Staubli VAL3: ForceData.pjx

--- ForceData.pjx ---
Parameters version=s8.15.3Cs9_BS3337 stackSize=5000 millimeterUnit=true
Data file=ForceData.dtx
Type name=tForce4Item path=Disk://LibTorque/template/Force4Item/Force4Item.pjx
Type name=tForce6Item path=Disk://LibTorque/template/Force6Item/Force6Item.pjx

--- ForceData.dtx ---
public tForce4Item tArm4Force{}
  [tp_80]
    num nMaxJnt4Force[4]
      [0] = 1029
      [1] = 254
      [2] = 833
      [3] = 15.2
    string sArmType
  [ts2_100]
    num nMaxJnt4Force[4]
      [0] = 570
      [1] = 255
      [2] = 789
      [3] = 15.6
    string sArmType
  [ts2_40]
    num nMaxJnt4Force[4]
      [0] = 570
      [1] = 255
      [2] = 789
      [3] = 15.6
    string sArmType
  [ts2_60]
    num nMaxJnt4Force[4]
      [0] = 570
      [1] = 255
      [2] = 789
      [3] = 15.6
    string sArmType
  [ts2_80]
    num nMaxJnt4Force[4]
      [0] = 570
      [1] = 255
      [2] = 789
      [3] = 15.6
    string sArmType
  [ts_20]
    num nMaxJnt4Force[4]
      [0] = 1029
      [1] = 137
      [2] = 789
      [3] = 15.6
    string sArmType
  [ts_40]
    num nMaxJnt4Force[4]
      [0] = 1029
      [1] = 137
      [2] = 789
      [3] = 15.6
    string sArmType
  [ts_60]
    num nMaxJnt4Force[4]
      [0] = 1029
      [1] = 137
      [2] = 789
      [3] = 15.6
    string sArmType
  [ts_80]
    num nMaxJnt4Force[4]
      [0] = 1029
      [1] = 137
      [2] = 789
      [3] = 15.6
    string sArmType
public tForce6Item tArm6Force{}
  [rx_160]
    num nMaxJnt6Force[6]
      [0] = 2660
      [1] = 2660
      [2] = 1128
      [3] = 570
      [4] = 248
      [5] = 153
    string sArmType
  [rx_160l]
    num nMaxJnt6Force[6]
      [0] = 2660
      [1] = 2660
      [2] = 1128
      [3] = 570
      [4] = 248
      [5] = 153
    string sArmType
  [tx2_140]
    num nMaxJnt6Force[6]
      [0] = 4280
      [1] = 4280
      [2] = 1128
      [3] = 570
      [4] = 255
      [5] = 86.4
    string sArmType
  [tx2_160]
    num nMaxJnt6Force[6]
      [0] = 4280
      [1] = 4280
      [2] = 1128
      [3] = 570
      [4] = 255
      [5] = 86.4
    string sArmType
  [tx2_160l]
    num nMaxJnt6Force[6]
      [0] = 4280
      [1] = 4280
      [2] = 1128
      [3] = 570
      [4] = 255
      [5] = 86.4
    string sArmType
  [tx2_200]
    num nMaxJnt6Force[6]
      [0] = 7840
      [1] = 7840
      [2] = 6207
      [3] = 3103
      [4] = 1383
      [5] = 1029
    string sArmType
  [tx2_200l]
    num nMaxJnt6Force[6]
      [0] = 7840
      [1] = 7840
      [2] = 6207
      [3] = 3103
      [4] = 1383
      [5] = 1029
    string sArmType
  [tx2_40]
    num nMaxJnt6Force[6]
      [0] = 197
      [1] = 197
      [2] = 60
      [3] = 60
      [4] = 22.4
      [5] = 13.6
    string sArmType
  [tx2_60]
    num nMaxJnt6Force[6]
      [0] = 560
      [1] = 560
      [2] = 197
      [3] = 60
      [4] = 25
      [5] = 25
    string sArmType
  [tx2_60l]
    num nMaxJnt6Force[6]
      [0] = 560
      [1] = 560
      [2] = 197
      [3] = 60
      [4] = 25
      [5] = 25
    string sArmType
  [tx2_90]
    num nMaxJnt6Force[6]
      [0] = 1128
      [1] = 1128
      [2] = 560
      [3] = 197
      [4] = 76.8
      [5] = 74
    string sArmType
  [tx2_90l]
    num nMaxJnt6Force[6]
      [0] = 1128
      [1] = 1128
      [2] = 560
      [3] = 197
      [4] = 76.8
      [5] = 74
    string sArmType
  [tx2_90xl]
    num nMaxJnt6Force[6]
      [0] = 1128
      [1] = 1128
      [2] = 560
      [3] = 197
      [4] = 56
      [5] = 74
    string sArmType
  [tx_200]
    num nMaxJnt6Force[6]
      [0] = 7840
      [1] = 7840
      [2] = 6207
      [3] = 3103
      [4] = 1383
      [5] = 1029
    string sArmType
  [tx_200l]
    num nMaxJnt6Force[6]
      [0] = 7840
      [1] = 7840
      [2] = 6207
      [3] = 3103
      [4] = 1383
      [5] = 1029
    string sArmType
  [tx_40]
    num nMaxJnt6Force[6]
      [0] = 197
      [1] = 197
      [2] = 75
      [3] = 75
      [4] = 28
      [5] = 17
    string sArmType
  [tx_60]
    num nMaxJnt6Force[6]
      [0] = 560
      [1] = 560
      [2] = 197
      [3] = 31.2
      [4] = 25
      [5] = 25
    string sArmType
  [tx_60l]
    num nMaxJnt6Force[6]
      [0] = 560
      [1] = 560
      [2] = 197
      [3] = 31.2
      [4] = 25
      [5] = 25
    string sArmType
  [tx_60xl]
    num nMaxJnt6Force[6]
      [0] = 560
      [1] = 560
      [2] = 197
      [3] = 31.2
      [4] = 25
      [5] = 25
    string sArmType
  [tx_90]
    num nMaxJnt6Force[6]
      [0] = 1128
      [1] = 1128
      [2] = 560
      [3] = 197
      [4] = 76.8
      [5] = 74
    string sArmType
  [tx_90l]
    num nMaxJnt6Force[6]
      [0] = 1128
      [1] = 1128
      [2] = 560
      [3] = 197
      [4] = 76.8
      [5] = 74
    string sArmType
  [tx_90xl]
    num nMaxJnt6Force[6]
      [0] = 1128
      [1] = 1128
      [2] = 560
      [3] = 197
      [4] = 76.8
      [5] = 74
    string sArmType
